(* IEC 61131-3 sources: IEC61131-3_ST_SCL_Mutation_Generator/tools/plcverif, 2 files *)

(* ---- M096.st ---- *)
FUNCTION_BLOCK DEC_TO_HEX
  VAR_INPUT
    DecimalValue : DINT;
  END_VAR
  VAR_OUTPUT
    HexString : STRING;
  END_VAR
  VAR
    i : INT;
    hexDigits : ARRAY [0..15] OF STRING := ['0', '1', '2', '3', '4', '5', '6', '7', '8', '9', 'A', 'B', 'C', 'D', 'E', 'F'];
    digitIndex : INT;
    hexDigit : STRING;
    significantDigitFound : BOOL := FALSE;
    digitValue : DINT;
    powerOfInteger : DINT;
  END_VAR

  HexString := '';

  IF DecimalValue = 0 THEN
      HexString := '0';
      RETURN;
  END_IF;

  significantDigitFound := FALSE;

  FOR digitIndex := 0 TO 7 DO

      powerOfInteger:=1;
      FOR i := 1 TO 7 - digitIndex DO
        powerOfInteger := powerOfInteger * 16;
      END_FOR;

      digitValue := DIV(DecimalValue, powerOfInteger) MOD 16;
      hexDigit := hexDigits[digitValue];

      IF NOT (hexDigit <> '0' OR significantDigitFound OR (7 - digitIndex) = 0) THEN (* MUTATED: COND_NEGATE *)
          significantDigitFound := TRUE;
          HexString := CONCAT(HexString, hexDigit);
      END_IF;

  END_FOR;
END_FUNCTION_BLOCK

(* ---- pump.st ---- *)
FUNCTION_BLOCK "PumpControl"
{ S7_Optimized_Access := 'TRUE' }
VERSION : 0.1
VAR_INPUT
HighLevelSensor : Bool; // True if water is dangerously high
LowLevelSensor : Bool; // True if tank is empty
ManualStop : Bool;
END_VAR

VAR_OUTPUT
MainPump : Bool;
BackupPump : Bool;
END_VAR

BEGIN
// Main Pump Logic
IF #HighLevelSensor AND NOT #ManualStop THEN
#MainPump := TRUE;
ELIF #LowLevelSensor OR #ManualStop THEN
#MainPump := FALSE;
END_IF;

// Safety Backup Pump Logic IF #HighLevelSensor AND #MainPump THEN #BackupPump := TRUE;
// Turns on if main pump isnt enough or failed ELIF #LowLevelSensor THEN #BackupPump := FALSE; END_IF;
END_FUNCTION_BLOCK
